FUNCTION_BLOCK EPUCK_MOTORS (* E-puck wheels speed determiner *)
  (* Standard: 61499-2; Classification: SIFB; ApplicationDomain: Robotics; Function: Actuator; Type: SIFB; Description: LEFT and RIGHT paces(-1000 to 1000) *)
  (* Version 1.0, 2026-10-22, Mauricio Martins Taques Filho, GASR/UDESC, Initial version *)
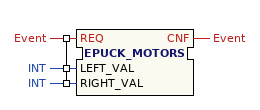
  EVENT_INPUT
    REQ WITH LEFT_VAL, RIGHT_VAL; (* Speed values *)
  END_EVENT
  EVENT_OUTPUT
    CNF; (* Set speeds *)
  END_EVENT
  VAR_INPUT
    LEFT_VAL : INT := 0; (* Left wheel paces *)
    RIGHT_VAL : INT := 0; (* Right wheel paces *)
  END_VAR
  SERVICE APPLICATION/RESOURCE
    SEQUENCE move_epuck
      APPLICATION.REQ(LEFT,RIGHT) -> APPLICATION.CNF();
    END_SEQUENCE
  END_SERVICE
END_FUNCTION_BLOCK
